FUNCTION_BLOCK FB_UpsConfigApply // EMS config/ups → UPS Holding 설정 쓰기
(* EMS가 내린 주기적·펄스 방전 설정을 UPS에 쓰고 되읽어 확인한다 (UPS 설정). 2026-11-02.
   기반 없음(신규).
   대상: H50~H61, H7, H10 (v2.51). 온도보상(H62~H64)은 스케일 확인 전이라 쓰지 않는다.
   2026-11-16 (명세 v2.14 CF-UPS-01): 간헐충전 H57~H61 추가. H58·H59는 H57이 1이면 전압(0.1 V), 2이면 SOC를
   같은 레지스터에 쓴다. EMS 4칸(전압 2, SOC 2) 중 기준에 맞는 2칸만 쓴다. 기준은 받은 값 → 보관값 → UPS 현재 H57 순.
   - 값 하나라도 범위 밖이면 그 UPS의 이번 설정 전체를 버린다 (BadConfig).
   - is_available=0인 필드와 현재 값이 같은 필드는 쓰지 않는다.
   - BAT Mode가 0(부동충전)일 때만 쓴다. 다른 운전 중이면 끝날 때까지 기다린다.
   - 쓰기 금지 상태에서 받은 설정은 적용하지 않고 버린다 (Disabled). 나중에 허용돼도 옛 값을 쓰지 않음.
   단위: 전류 A → 0.1A, 시간 분·초, 횟수 Cycle. EMS 쪽 단위는 확인 필요.
   2026-11-25 (명세 v2.51 CF-UPS-01): H7 부동 충전 전압·H10 충전 전류 추가 (칸 12·13, 값 × 10). 주소가 이어지지 않아
   칸 → 주소를 ITEM_ADDR 표로 찾는다. 범위: H7 0 초과 UPS_CFG_MAX_VOLTAGE_V 이하, H10 0 초과 UPS_CFG_MAX_CURRENT_A 이하.
   2026-11-23: M_Load가 VAR_IN_OUT(iq_stDesired)을 직접 읽던 것을 입력으로 넘김 (컴파일 경고 제거, 동작 같음)
   2026-11-05 (명세 CF-UPS-02·03): 받은 설정을 보관값(iq_stDesired, GVL_PERSIST)에 남기고,
   i_tRecheck마다 UPS 값을 되읽어 보관값과 다르면 다시 쓴다 (UPS 재기동·PMS 재시작·통신 복구 후 복구).
   UPS 고장(i_bUpsFault)·e-stop 중에는 쓰지 않는다. 2026-11-17: 쓰기 요청(20)·되읽기(30) 단계에서도 매 스캔 다시 보고,
   고장·e-stop·부동충전 아님·데이터 무효면 10단계로 돌아가 기다린다 (실패로 세지 않음). 쓰기가 i_nMaxFail회 연속 실패하면 q_bMismatch를 켜고
   새 설정을 받을 때까지 복구를 멈춘다. *)
VAR_INPUT
	i_bEnable : BOOL; // 장비 쓰기 허용
	i_nRxCount : UDINT; // config/ups 수신 누계
	i_stConfig : ST_UpsConfig_Rx; // 이 UPS의 수신 설정
	i_stState : ST_UpsState; // 장비 상태
	i_stRaw : ST_UpsRaw; // 되읽기용 원본
	i_ipUps : I_Ups; // 쓰기 대상
	i_tTimeout : TIME := T#10S; // 주소 하나의 쓰기·되읽기 제한 시간
	i_bUpsFault : BOOL; // UPS 고장 있음 (보고 Status b6). 켜져 있으면 쓰지 않음
	i_tRecheck : TIME := T#10S; // 보관값과 UPS 값을 비교하는 주기
	i_nMaxFail : UINT := 3; // 연속 실패 허용 횟수. 넘으면 q_bMismatch
END_VAR
VAR_IN_OUT
	iq_stDesired : ST_UpsDesiredSet; // 맞춰 둘 설정 보관값 (GVL_PERSIST.g_astUpsDesired[n])
END_VAR
VAR_OUTPUT
	q_bBusy : BOOL; // 적용 중
	q_eResult : E_UpsResult; // 마지막 적용 결과
	q_nErrorAddress : UINT; // 실패한 H 주소. 0 = 없음
	q_nAppliedRx : UDINT; // 마지막으로 처리한 수신 누계
	q_nWriteCount : UDINT; // 적용한 주소 수 누계
	q_bDesiredChanged : BOOL; // 이 스캔에 보관값을 바꿈 (PERSISTENT 바로 저장 요청)
	q_bMismatch : BOOL; // 설정 불일치 알람: 연속 i_nMaxFail회 실패. 새 설정을 받으면 풀림
	q_nRecoverCount : UDINT; // 복구로 다시 쓴 주소 수 누계
END_VAR
VAR CONSTANT
	ITEM_COUNT : UINT := 14;
	ITEM_ADDR : ARRAY[0..ITEM_COUNT-1] OF UINT := [50, 51, 52, 53, 54, 55, 56, 57, 58, 59, 60, 61, 7, 10]; // 칸 → H 주소. H50~H61, H7, H10 (명세 v2.51)
END_VAR
VAR
	_nStep : UINT;
	_nItem : UINT;
	_nLastRx : UDINT;
	_bBad : BOOL;
	_awTarget : ARRAY[0..ITEM_COUNT-1] OF WORD; // 쓸 값
	_abUse : ARRAY[0..ITEM_COUNT-1] OF BOOL;
	_tonTimeout : TON;
	_tonRecheck : TON; // 비교 주기
	_bRecover : BOOL; // 지금 진행 중인 쓰기가 복구인지 (수신이 아니라)
	_nFail : UINT; // 연속 실패 횟수
	_nCheck : UINT;
END_VAR

_tonTimeout(IN:=_nStep=20 OR _nStep=30, PT:=i_tTimeout);
_tonRecheck(IN:=_nStep=0 AND NOT _tonRecheck.Q, PT:=i_tRecheck);
q_bDesiredChanged:=FALSE;

CASE _nStep OF
	0: // 새 설정 대기
		q_bBusy:=FALSE;
		IF i_nRxCount<>_nLastRx THEN
			_nLastRx:=i_nRxCount;
			q_nErrorAddress:=0;
			IF NOT i_bEnable OR i_ipUps=0 THEN
				q_eResult:=E_UpsResult.Disabled;
				q_nAppliedRx:=_nLastRx;
			ELSE
				M_Load(i_bSavedMode:=iq_stDesired.bValid AND iq_stDesired.abUse[7], i_wSavedMode:=iq_stDesired.awValue[7]);
				IF _bBad THEN
					q_eResult:=E_UpsResult.BadConfig;
					q_nAppliedRx:=_nLastRx;
				ELSE
					// 받은 설정을 보관값으로 남김 (CF-UPS-02)
					iq_stDesired.abUse:=_abUse;
					iq_stDesired.awValue:=_awTarget;
					iq_stDesired.nRxCount:=_nLastRx;
					iq_stDesired.bValid:=TRUE;
					q_bDesiredChanged:=TRUE;
					q_bMismatch:=FALSE;
					_nFail:=0;
					_bRecover:=FALSE;
					q_bBusy:=TRUE;
					q_eResult:=E_UpsResult.Busy;
					_nItem:=0;
					_nStep:=10;
				END_IF
			END_IF
		ELSIF _tonRecheck.Q AND iq_stDesired.bValid AND i_bEnable AND i_ipUps<>0 AND NOT q_bMismatch AND i_stState.bValid THEN
			// 복구 (CF-UPS-03): 보관값과 UPS 값이 다른 칸이 있으면 다시 쓴다
			_abUse:=iq_stDesired.abUse;
			_awTarget:=iq_stDesired.awValue;
			_bRecover:=FALSE;
			FOR _nCheck:=0 TO ITEM_COUNT-1 DO
				IF _abUse[_nCheck] AND i_stRaw.awParam[ITEM_ADDR[_nCheck]]<>_awTarget[_nCheck] THEN
					_bRecover:=TRUE;
				END_IF
			END_FOR
			IF _bRecover THEN
				q_nErrorAddress:=0;
				q_bBusy:=TRUE;
				q_eResult:=E_UpsResult.Busy;
				_nItem:=0;
				_nStep:=10;
			END_IF
		END_IF

	10: // 부동충전 상태에서만 진행
		IF NOT i_bEnable THEN
			q_eResult:=E_UpsResult.Disabled;
			q_nAppliedRx:=_nLastRx;
			_nStep:=0;
		ELSIF i_stState.bValid AND i_stState.nBatMode=0 AND NOT i_bUpsFault AND NOT i_stState.bEmergencyStop THEN
			WHILE _nItem<ITEM_COUNT DO
				IF _abUse[_nItem] AND i_stRaw.awParam[ITEM_ADDR[_nItem]]<>_awTarget[_nItem] THEN EXIT; END_IF
				_nItem:=_nItem+1;
			END_WHILE
			IF _nItem>=ITEM_COUNT THEN
				q_eResult:=E_UpsResult.Accepted;
				q_nAppliedRx:=_nLastRx;
				_nFail:=0;
				_bRecover:=FALSE;
				_nStep:=0;
			ELSE
				_nStep:=20;
			END_IF
		END_IF

	20: // 쓰기 요청
		IF NOT i_bEnable THEN
			q_eResult:=E_UpsResult.Disabled;
			q_nAppliedRx:=_nLastRx;
			_nStep:=0;
		ELSIF i_bUpsFault OR i_stState.bEmergencyStop OR NOT i_stState.bValid OR i_stState.nBatMode<>0 THEN
			_nStep:=10; // 2026-11-17: 기다리는 동안 고장·e-stop 등이 생김 → 쓰지 않고 10단계에서 기다림
		ELSIF i_ipUps.M_SetParameter(UINT_TO_WORD(ITEM_ADDR[_nItem]),_awTarget[_nItem]) THEN
			_nStep:=30;
		ELSIF _tonTimeout.Q THEN
			_nStep:=900;
		END_IF

	30: // 되읽기 확인
		IF i_bUpsFault OR i_stState.bEmergencyStop THEN
			_nStep:=10; // 2026-11-17: 드라이버가 고장·e-stop으로 쓰기를 뺐을 수 있음 → 실패로 세지 않고 다시 기다림
		ELSIF i_stRaw.awParam[ITEM_ADDR[_nItem]]=_awTarget[_nItem] THEN
			q_nWriteCount:=q_nWriteCount+1;
			IF _bRecover THEN q_nRecoverCount:=q_nRecoverCount+1; END_IF
			_nItem:=_nItem+1;
			_nStep:=10;
		ELSIF _tonTimeout.Q THEN
			_nStep:=900;
		END_IF

	900: // 실패. 남은 주소는 쓰지 않음
		q_eResult:=E_UpsResult.CommUnavailable;
		q_nErrorAddress:=ITEM_ADDR[_nItem];
		q_nAppliedRx:=_nLastRx;
		_nFail:=_nFail+1;
		IF _nFail>=i_nMaxFail THEN q_bMismatch:=TRUE; END_IF // 반복을 멈추고 알람
		_bRecover:=FALSE;
		_nStep:=0;
END_CASE

METHOD PRIVATE M_Load
VAR_INPUT
	i_bSavedMode : BOOL; // 보관값에 간헐충전 기준(H57)이 있음 (iq_stDesired.bValid AND abUse[7])
	i_wSavedMode : WORD; // 그 기준 값 (iq_stDesired.awValue[7])
END_VAR
VAR
	nMode : UDINT; // 간헐충전 기준 0 끔 / 1 전압 / 2 SOC (H57)
	bStartAv : BOOL; // 기준에 맞는 시작 칸을 받음
	bEndAv : BOOL; // 기준에 맞는 종료 칸을 받음
	rStart : REAL;
	rEnd : REAL;
	rScale : REAL; // 레지스터 배율 (전압 10, SOC GVL_PARAM.UPS_CFG_SOC_SCALE)
	rMax : REAL; // 상한 (전압 UPS_CFG_MAX_VOLTAGE_V, SOC 100)
END_VAR
_bBad:=FALSE;
_abUse[0]:=i_stConfig.PeriodicTrickleDischargeSetCurrent.is_available<>0;
IF _abUse[0] THEN
	IF i_stConfig.PeriodicTrickleDischargeSetCurrent.value>0.0 AND i_stConfig.PeriodicTrickleDischargeSetCurrent.value<=GVL_PARAM.UPS_CFG_MAX_CURRENT_A THEN
		_awTarget[0]:=REAL_TO_WORD(i_stConfig.PeriodicTrickleDischargeSetCurrent.value*10.0);
	ELSE _bBad:=TRUE; q_nErrorAddress:=50; END_IF
END_IF
_abUse[1]:=i_stConfig.PeriodicTrickleDischargeSetTime.is_available<>0;
IF _abUse[1] THEN
	IF i_stConfig.PeriodicTrickleDischargeSetTime.value>0 AND i_stConfig.PeriodicTrickleDischargeSetTime.value<=GVL_PARAM.UPS_CFG_MAX_MINUTES THEN
		_awTarget[1]:=UDINT_TO_WORD(i_stConfig.PeriodicTrickleDischargeSetTime.value);
	ELSE _bBad:=TRUE; q_nErrorAddress:=51; END_IF
END_IF
_abUse[2]:=i_stConfig.PulseDischargeSetCurrent.is_available<>0;
IF _abUse[2] THEN
	IF i_stConfig.PulseDischargeSetCurrent.value>0.0 AND i_stConfig.PulseDischargeSetCurrent.value<=GVL_PARAM.UPS_CFG_MAX_CURRENT_A THEN
		_awTarget[2]:=REAL_TO_WORD(i_stConfig.PulseDischargeSetCurrent.value*10.0);
	ELSE _bBad:=TRUE; q_nErrorAddress:=52; END_IF
END_IF
_abUse[3]:=i_stConfig.PulseChargeSetCurrent.is_available<>0;
IF _abUse[3] THEN
	IF i_stConfig.PulseChargeSetCurrent.value>0.0 AND i_stConfig.PulseChargeSetCurrent.value<=GVL_PARAM.UPS_CFG_MAX_CURRENT_A THEN
		_awTarget[3]:=REAL_TO_WORD(i_stConfig.PulseChargeSetCurrent.value*10.0);
	ELSE _bBad:=TRUE; q_nErrorAddress:=53; END_IF
END_IF
_abUse[4]:=i_stConfig.PulseDischargeSetTime.is_available<>0;
IF _abUse[4] THEN
	IF i_stConfig.PulseDischargeSetTime.value>0 AND i_stConfig.PulseDischargeSetTime.value<=GVL_PARAM.UPS_CFG_MAX_SECONDS THEN
		_awTarget[4]:=UDINT_TO_WORD(i_stConfig.PulseDischargeSetTime.value);
	ELSE _bBad:=TRUE; q_nErrorAddress:=54; END_IF
END_IF
_abUse[5]:=i_stConfig.PulseChargeSetTime.is_available<>0;
IF _abUse[5] THEN
	IF i_stConfig.PulseChargeSetTime.value>0 AND i_stConfig.PulseChargeSetTime.value<=GVL_PARAM.UPS_CFG_MAX_SECONDS THEN
		_awTarget[5]:=UDINT_TO_WORD(i_stConfig.PulseChargeSetTime.value);
	ELSE _bBad:=TRUE; q_nErrorAddress:=55; END_IF
END_IF
_abUse[6]:=i_stConfig.PulseChargeDischargeSetCycle.is_available<>0;
IF _abUse[6] THEN
	IF i_stConfig.PulseChargeDischargeSetCycle.value>0 AND i_stConfig.PulseChargeDischargeSetCycle.value<=GVL_PARAM.UPS_CFG_MAX_CYCLES THEN
		_awTarget[6]:=UDINT_TO_WORD(i_stConfig.PulseChargeDischargeSetCycle.value);
	ELSE _bBad:=TRUE; q_nErrorAddress:=56; END_IF
END_IF
// H57~H61 간헐충전 (명세 v2.14 CF-UPS-01). H58·H59는 H57 기준에 따라 전압 또는 SOC
_abUse[7]:=i_stConfig.TrickleChargeSetParameter.is_available<>0;
IF _abUse[7] THEN
	IF i_stConfig.TrickleChargeSetParameter.value<=2 THEN
		nMode:=i_stConfig.TrickleChargeSetParameter.value;
		_awTarget[7]:=UDINT_TO_WORD(nMode);
	ELSE _bBad:=TRUE; q_nErrorAddress:=57; END_IF
ELSIF i_bSavedMode THEN
	nMode:=WORD_TO_UDINT(i_wSavedMode);
ELSE
	nMode:=WORD_TO_UDINT(i_stRaw.awParam[57]);
END_IF
_abUse[8]:=FALSE;
_abUse[9]:=FALSE;
bStartAv:=FALSE;
bEndAv:=FALSE;
IF nMode=1 THEN
	bStartAv:=i_stConfig.TrickleChargeSetStartVoltage.is_available<>0;
	bEndAv:=i_stConfig.TrickleChargeSetEndVoltage.is_available<>0;
	rStart:=i_stConfig.TrickleChargeSetStartVoltage.value;
	rEnd:=i_stConfig.TrickleChargeSetEndVoltage.value;
	rScale:=10.0;
	rMax:=GVL_PARAM.UPS_CFG_MAX_VOLTAGE_V;
ELSIF nMode=2 THEN
	bStartAv:=i_stConfig.TrickleChargeSetStartSoc.is_available<>0;
	bEndAv:=i_stConfig.TrickleChargeSetEndSoc.is_available<>0;
	rStart:=i_stConfig.TrickleChargeSetStartSoc.value;
	rEnd:=i_stConfig.TrickleChargeSetEndSoc.value;
	rScale:=GVL_PARAM.UPS_CFG_SOC_SCALE;
	rMax:=100.0;
END_IF
IF nMode=1 OR nMode=2 THEN
	IF _abUse[7] AND NOT (bStartAv AND bEndAv) THEN
		_bBad:=TRUE; q_nErrorAddress:=58; // 기준을 바꿀 때는 시작·종료를 같이 받아야 함
	ELSE
		IF bStartAv AND bEndAv AND rStart>=rEnd THEN _bBad:=TRUE; q_nErrorAddress:=58; END_IF
		IF bStartAv THEN
			IF rStart>0.0 AND rStart<=rMax THEN _abUse[8]:=TRUE; _awTarget[8]:=REAL_TO_WORD(rStart*rScale);
			ELSE _bBad:=TRUE; q_nErrorAddress:=58; END_IF
		END_IF
		IF bEndAv THEN
			IF rEnd>0.0 AND rEnd<=rMax THEN _abUse[9]:=TRUE; _awTarget[9]:=REAL_TO_WORD(rEnd*rScale);
			ELSE _bBad:=TRUE; q_nErrorAddress:=59; END_IF
		END_IF
	END_IF
END_IF
_abUse[10]:=i_stConfig.TrickleChargeSetStartTime.is_available<>0; // EMS 이름은 StartTime, 맵 H60은 간헐충전 종료시간 (분)
IF _abUse[10] THEN
	IF i_stConfig.TrickleChargeSetStartTime.value>0 AND i_stConfig.TrickleChargeSetStartTime.value<=GVL_PARAM.UPS_CFG_MAX_TRICKLE_MINUTES THEN
		_awTarget[10]:=UDINT_TO_WORD(i_stConfig.TrickleChargeSetStartTime.value);
	ELSE _bBad:=TRUE; q_nErrorAddress:=60; END_IF
END_IF
_abUse[11]:=i_stConfig.TrickleChargeSetReStartDay.is_available<>0;
IF _abUse[11] THEN
	IF i_stConfig.TrickleChargeSetReStartDay.value>0 AND i_stConfig.TrickleChargeSetReStartDay.value<=GVL_PARAM.UPS_CFG_MAX_DAYS THEN
		_awTarget[11]:=UDINT_TO_WORD(i_stConfig.TrickleChargeSetReStartDay.value);
	ELSE _bBad:=TRUE; q_nErrorAddress:=61; END_IF
END_IF
// H7 부동 충전 전압·H10 충전 전류 (명세 v2.51 CF-UPS-01). 값 × 10
_abUse[12]:=i_stConfig.FloatChargeSetVoltage.is_available<>0;
IF _abUse[12] THEN
	IF i_stConfig.FloatChargeSetVoltage.value>0.0 AND i_stConfig.FloatChargeSetVoltage.value<=GVL_PARAM.UPS_CFG_MAX_VOLTAGE_V THEN
		_awTarget[12]:=REAL_TO_WORD(i_stConfig.FloatChargeSetVoltage.value*10.0);
	ELSE _bBad:=TRUE; q_nErrorAddress:=7; END_IF
END_IF
_abUse[13]:=i_stConfig.ChargeSetCurrentLimit.is_available<>0;
IF _abUse[13] THEN
	IF i_stConfig.ChargeSetCurrentLimit.value>0.0 AND i_stConfig.ChargeSetCurrentLimit.value<=GVL_PARAM.UPS_CFG_MAX_CURRENT_A THEN
		_awTarget[13]:=REAL_TO_WORD(i_stConfig.ChargeSetCurrentLimit.value*10.0);
	ELSE _bBad:=TRUE; q_nErrorAddress:=10; END_IF
END_IF
END_METHOD

END_FUNCTION_BLOCK

(* stored: Version 1.1.0.1, ProductVersion 3.1.4024.15
   POU FB_UpsConfigApply: Id {4e08e92f-3455-48e2-9428-4f5d2d75fec4}, SpecialFunc None
   Method M_Load: Id {00b4605e-ed77-4b5f-9061-112fb14dbe73} *)
